(* IEC 61131-3 sources: Gen-AI/docs/member2_validation/codesys_release_v1.1/C01_undeclared, 1 file *)

(* ---- source.st ---- *)
FUNCTION_BLOCK FB_AgentProbeUndeclared
VAR_OUTPUT
 y : BOOL;
END_VAR
y := AgentSignalNotDeclared_6E79B1;
END_FUNCTION_BLOCK
